// TwinCAT 3 PLC project PLC_ReadWriteCsvFile
// ProgramVersion: 3.1.4026.30
// libraries:
//   Tc2_Standard, * (Beckhoff Automation GmbH)
//   Tc2_System, * (Beckhoff Automation GmbH)
//   Tc2_Utilities, * (Beckhoff Automation GmbH)
//   Tc3_Mc3FluidPower, * (Beckhoff Automation GmbH)
//   Tc3_Mc3FluidPower_Preview, * (Beckhoff Automation GmbH)
//   Tc3_Module, * (Beckhoff Automation GmbH)
// project tree:
//   / PlcTask.TcTTO
//   POUs/ MAIN.TcPOU
// real-time tasks:
//   TASK PlcTask: cycle T#10ms, priority 20, ADS port 350

CONFIGURATION PLC_ReadWriteCsvFile
    RESOURCE PLC ON TwinCAT3
        TASK PlcTask(INTERVAL := T#10ms, PRIORITY := 20);
        PROGRAM MAIN WITH PlcTask : MAIN;
    END_RESOURCE
END_CONFIGURATION

// ---- POUs/MAIN.TcPOU
// Valve Characteristic Curve - Read/Write CSV sample
// Shows persisting valve characteristic curve data (SpoolPosition/Velocity points) to and from
// CSV files with MC_ValveCharacteristicCurve_WriteToCsv / _ReadFromCsv.
// Operation: set bStartWrite := TRUE to write, bStartRead := TRUE to read; bUseComma selects the CSV field separator.
PROGRAM MAIN
VAR  
	/// the filepath '/temp/ValveCharacteristicCurve.csv' requests the folder 'temp' in C:\
  
    (* Configuration *)
    bUseComma : BOOL;
    
    (* Controls *)
    bStartWrite : BOOL;
    bStartRead  : BOOL;
    
    fbRead  : MC_ValveCharacteristicCurve_ReadFromCsv;
    fbWrite : MC_ValveCharacteristicCurve_WriteToCsv;
    aWriteData : ARRAY[1..5] OF ValveCharacteristicPoint := [(Velocity:=-1.0, SpoolPosition:=-1.0), (Velocity:=-0.8, SpoolPosition:=-0.5), (Velocity:=0.0, SpoolPosition:=0.0), (Velocity:=0.4, SpoolPosition:=0.5), (Velocity:=0.8, SpoolPosition:=1.0)];
END_VAR

(* Set CSV field separator to ';' (16#3B) for comma decimals, or ',' (16#2C) otherwise *)
IF bUseComma THEN
	DEFAULT_CSV_FIELD_SEP := 16#2C; (* Comma *)
ELSE
    DEFAULT_CSV_FIELD_SEP := 16#3B; (* Semicolon *)
END_IF

IF bStartWrite THEN
    bStartWrite:=FALSE;
    fbWrite.Write:=TRUE;
    fbWrite.FilePath:='/temp/ValveCharacteristicCurve.csv';
END_IF

IF bStartRead THEN
    bStartRead:=FALSE;
    fbRead.Read:=TRUE;
    fbRead.FilePath:='/temp/ValveCharacteristicCurve.csv';
END_IF

fbWrite(DataPoints:=aWriteData);
fbRead();

END_PROGRAM
